DATA_BLOCK "GDB_ProfileIntegration"
{ S7_Optimized_Access := 'TRUE' }
VERSION : 0.1
NON_RETAIN
VAR
    Owner : DInt;
    Enabled : Bool;
    StepNo : DInt;
    Branch : DInt;
    TimeClass : DInt;
    Expected : Time;
    Finish : Bool;
    ForceLateTimeout : Bool;
    RequestSeq : UDInt;
    AckSeq {ExternalWritable := 'False'} : UDInt;
END_VAR
BEGIN
END_DATA_BLOCK
